SUBAPPLICATION Uebung_136b (* Übung zu STRING über CAN senden (bis 8 Zeichen), Text vom VT *)
  (* Standard: 61499-2; Description: Copyright (c) 2026 Meisterschulen am Ostbahnhof This program and the accompanying materials are made available under the terms of the Eclipse Public License 2.0 which is available at https://www.eclipse.org/legal/epl-2.0/ SPDX-License-Identifier: EPL-2.0 *)
  (* Version 1.0, 2026-11-14, Franz Höpfinger, Meisterschulen am Ostbahnhof, initial API and implementation and/or initial documentation *)
  PACKAGE Uebungen;
  IMPORT Uebungen::const::UT::DefaultPool::InputString_S1;
  IMPORT Uebungen::const::Uebung_120_129::Filter::ADD_ALL_PASS;
  IMPORT Uebungen::const::Uebung_120_129::Filter::FLT_ALL_PASS;
  IMPORT isobus::pgn::ADDRESS::GLOBAL_A;
  IMPORT isobus::pgn::ISOUSERHOME_e::thisMember;
  IMPORT isobus::pgn::ISO_CAN_NODE::NODE1;
  IMPORT isobus::pgn::const::PgnDef::PGN_PDU1_PropA;
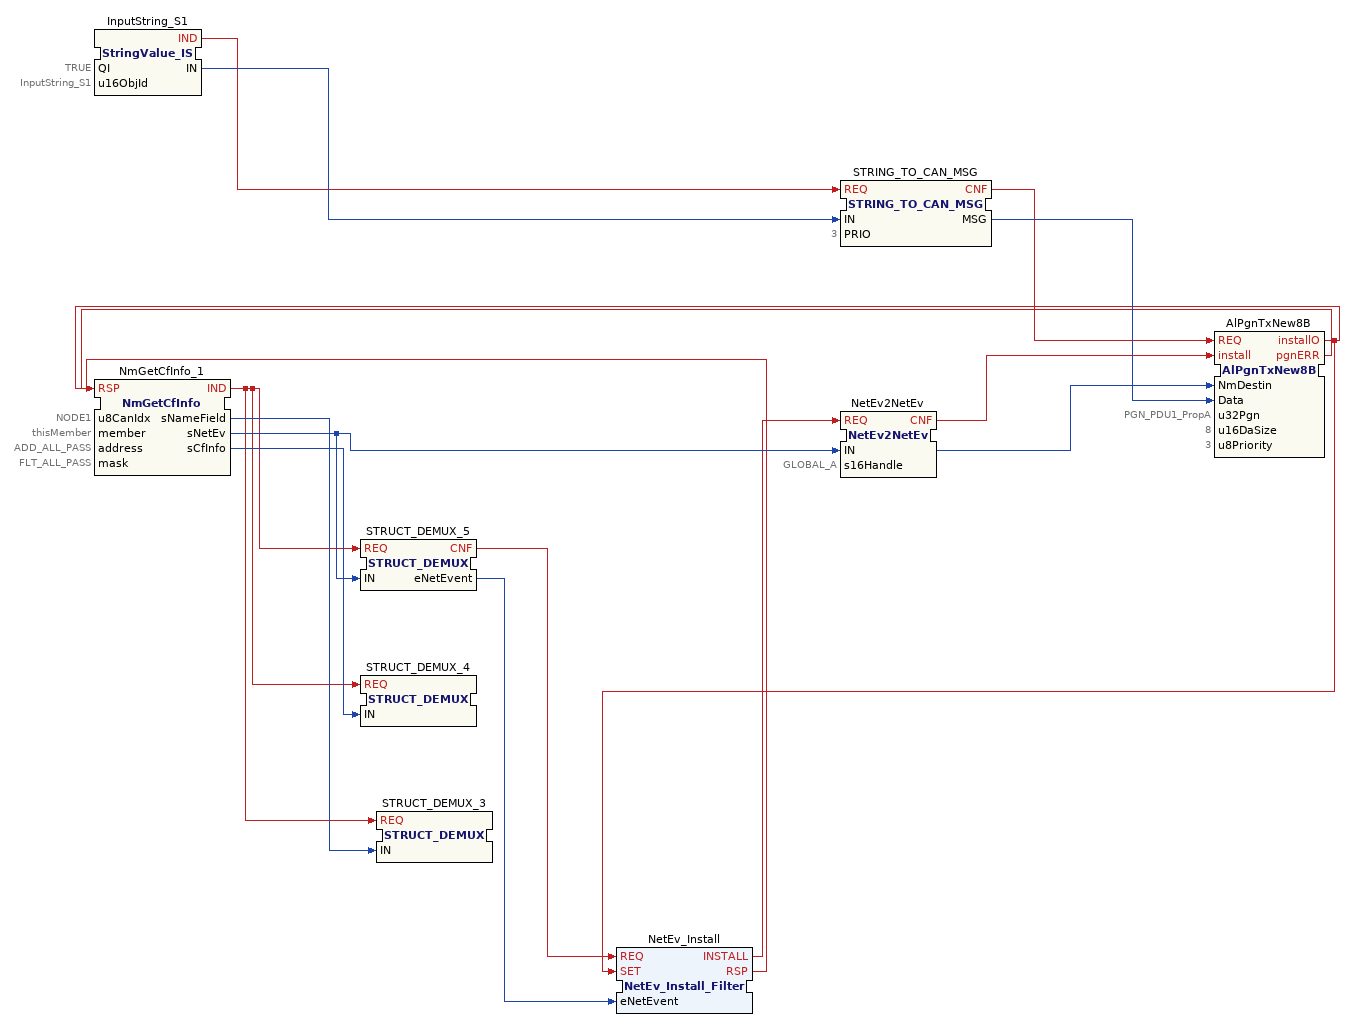
  FBS
    STRUCT_DEMUX_3 : eclipse4diac::convert::STRUCT_DEMUX; {SET_ATTRIBUTE(StructuredType, isobus::pgn::NAMEFIELD_T)}
    NmGetCfInfo_1 : isobus::pgn::NmGetCfInfo(u8CanIdx := NODE1, member := thisMember, address := ADD_ALL_PASS, mask := FLT_ALL_PASS);
    STRUCT_DEMUX_4 : eclipse4diac::convert::STRUCT_DEMUX; {SET_ATTRIBUTE(StructuredType, isobus::pgn::CF_INFO_T)}
    STRUCT_DEMUX_5 : eclipse4diac::convert::STRUCT_DEMUX; {SET_ATTRIBUTE(StructuredType, isobus::pgn::ISONETEVENT_T)}
    NetEv2NetEv : isobus::pgn::NetEv2NetEv(s16Handle := GLOBAL_A);
    STRING_TO_CAN_MSG : isobus::pgn::STRING_TO_CAN_MSG(PRIO := 3);
    AlPgnTxNew8B : isobus::pgn::tx::AlPgnTxNew8B(u32Pgn := PGN_PDU1_PropA, u16DaSize := 8, u8Priority := 3);
    InputString_S1 : isobus::UT::io::StringValue::StringValue_IS(QI := TRUE, u16ObjId := InputString_S1);
  END_FBS
  SUBAPPS
    NetEv_Install : MyLib::sys::NetEv_Install_Filter;
  END_SUBAPPS
  EVENT_CONNECTIONS
    NmGetCfInfo_1.IND TO STRUCT_DEMUX_3.REQ;
    NmGetCfInfo_1.IND TO STRUCT_DEMUX_4.REQ;
    NmGetCfInfo_1.IND TO STRUCT_DEMUX_5.REQ;
    InputString_S1.IND TO STRING_TO_CAN_MSG.REQ;
    STRING_TO_CAN_MSG.CNF TO AlPgnTxNew8B.REQ;
    NetEv2NetEv.CNF TO AlPgnTxNew8B.install;
    AlPgnTxNew8B.installO TO NmGetCfInfo_1.RSP;
    AlPgnTxNew8B.pgnERR TO NmGetCfInfo_1.RSP;
    STRUCT_DEMUX_5.CNF TO NetEv_Install.REQ;
    NetEv_Install.INSTALL TO NetEv2NetEv.REQ;
    NetEv_Install.RSP TO NmGetCfInfo_1.RSP;
    AlPgnTxNew8B.installO TO NetEv_Install.SET;
  END_CONNECTIONS
  DATA_CONNECTIONS
    NmGetCfInfo_1.sNameField TO STRUCT_DEMUX_3.IN;
    NmGetCfInfo_1.sNetEv TO STRUCT_DEMUX_5.IN;
    NmGetCfInfo_1.sCfInfo TO STRUCT_DEMUX_4.IN;
    NmGetCfInfo_1.sNetEv TO NetEv2NetEv.IN;
    InputString_S1.IN TO STRING_TO_CAN_MSG.IN;
    NetEv2NetEv. TO AlPgnTxNew8B.NmDestin;
    STRING_TO_CAN_MSG.MSG TO AlPgnTxNew8B.Data;
    STRUCT_DEMUX_5.eNetEvent TO NetEv_Install.eNetEvent;
  END_CONNECTIONS
END_SUBAPPLICATION
